FUNCTION_BLOCK SENSOR_HISTORICAL_DB_WRITER
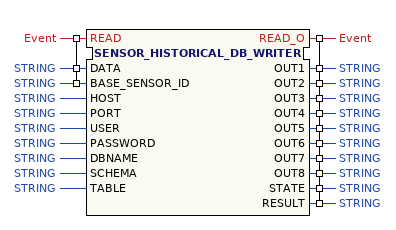
  EVENT_INPUT
    READ WITH DATA, BASE_SENSOR_ID;
  END_EVENT
  EVENT_OUTPUT
    READ_O WITH OUT1, OUT2, OUT3, OUT4, OUT5, OUT6, OUT7, OUT8, STATE, RESULT;
  END_EVENT
  VAR_INPUT
    DATA : STRING;
    BASE_SENSOR_ID : STRING;
    HOST : STRING;
    PORT : STRING;
    USER : STRING;
    PASSWORD : STRING;
    DBNAME : STRING;
    SCHEMA : STRING;
    TABLE : STRING;
  END_VAR
  VAR_OUTPUT
    OUT1 : STRING;
    OUT2 : STRING;
    OUT3 : STRING;
    OUT4 : STRING;
    OUT5 : STRING;
    OUT6 : STRING;
    OUT7 : STRING;
    OUT8 : STRING;
    STATE : STRING;
    RESULT : STRING;
  END_VAR
END_FUNCTION_BLOCK
